(* IEC 61131-3 sources: guidance-for-physical-ai-production-designer-on-aws/source/plan2cell/crates/plan2cell/tests/fixtures/deploy_check/welding_cell_2_small/plc/codesys/head/GVL, 1 file *)

(* ---- GVL_Cell.st ---- *)
(*
 * GVL_Cell - generated by bt2plc 0.1.0 - DO NOT EDIT
 * Plan   : bt_1792076124_welding_cell_2_small (cell welding_cell_2_small)
 * Grants : planned ticket order
 * IL01   : R1#1 W03 > R2#2 W14 > R1#3 W06 > R2#4 W10 > R1#5 ROBOT1_S04 > R2#6 W12 > R1#7 W05 > R2#8 ROBOT2_S07 > R1#9 ROBOT1_S08 > R2#10 W07 > R1#11 HOME
 * IL02   : R2#1 W15 > R1#2 W02 > R2#3 W13 > R1#4 W01 > R2#5 W11 > R1#6 W04 > R2#7 ROBOT2_S06 > R1#8 W08 > R2#9 W09 > R1#10 ROBOT1_S09 > R2#11 HOME
 *)
{attribute 'qualified_only'}
VAR_GLOBAL CONSTANT
    (* ========================================================================
       DIMENSIONS (array bounds are literals; *_DIM >= 1)
       ======================================================================== *)
    N_ROBOTS                : INT := 2;
    N_ZONES                 : INT := 2;
    N_OPS                   : INT := 22;
    N_PREDS                 : INT := 0;

    (* ========================================================================
       PROTOCOL / TIMING
       ======================================================================== *)
    PLAN_ID                 : WORD := WORD#16#4F80;             (* fold of the plan fingerprint *)
    PROD_FOLGE              : WORD := WORD#11;                  (* default production Folge *)
    HOME_FOLGE              : WORD := WORD#125;                 (* blind homing *)
    JOB_NUMBER_BYTE         : BOOL := FALSE;                    (* FALSE: WORD LE bytes 2-3, TRUE: byte 2 *)
    PROFILE_VW              : BOOL := FALSE;                    (* TRUE: VW KS24 signal map and Folge handshake instead of the simulator telegram *)
    GRANT_POLICY            : E_GrantPolicy := E_GrantPolicy.GP_PLANNED;
    HOME_SEQUENTIAL         : BOOL := TRUE;
    AUTO_RUN                : BOOL := TRUE;                     (* start the next cycle automatically *)
    STEP_BYTE               : INT := 4;                         (* robot -> PLC, WORD LE op index *)
    REQ_BYTE                : INT := 28;                        (* robot -> PLC, DWORD LE zone requests *)
    GRANT_BYTE              : INT := 12;                        (* PLC -> robot, DWORD LE zone grants *)
    PLAN_ID_BYTE            : INT := 4;                         (* PLC -> robot, WORD LE plan id *)
    PERMIT_MASK             : DWORD := DWORD#16#80000000;       (* bit 31: permit predecessors *)
    T_RESET_PULSE           : TIME := T#1S;
    T_START_PULSE           : TIME := T#500MS;
    T_STOP_PULSE            : TIME := T#1S;
    T_HANDSHAKE             : TIME := T#5S;
    T_BRINGUP_LIMIT         : TIME := T#1M;                     (* safety enable: PROFINET connection set-up *)
    T_MISMATCH_DEBOUNCE     : TIME := T#200MS;
    T_STOP_DEBOUNCE         : TIME := T#200MS;                  (* job running: ProgRunning and ProgFinished low this long = robot stopped *)
    T_CYCLE_PAUSE           : TIME := T#2S;
    T_START_LIMIT           : TIME := T#15S;
    T_ABORT_LIMIT           : TIME := T#10S;
    T_HOME_LIMIT            : TIME := T#15S500MS;

    (* ========================================================================
       VW KS24 SIGNAL INDICES (used when PROFILE_VW; $IN/$OUT index, 1-based)
       ======================================================================== *)
    VW_READY_OUT            : INT := 9;                         (* O_R_Bereit *)
    VW_RK100_OUT            : INT := 10;                        (* O_R_RK100 safety circuit *)
    VW_AUTO_OUT             : INT := 12;                        (* O_R_Auto *)
    VW_ESTOP_OUT            : INT := 13;                        (* O_R_Notaus *)
    VW_END_OUT              : INT := 14;                        (* O_R_F_ENDE / LPKT *)
    VW_PF0_OUT              : INT := 15;                        (* O_R_PFO home position *)
    VW_STEP_OUT             : INT := 97;                        (* P_PktNr_SPS op index (16 bits) *)
    VW_REL_OUT              : INT := 41;                        (* interlock releases A41-56 *)
    VW_REQ_OUT              : INT := 81;                        (* interlock requests A81-96 *)
    VW_ERR_OUT              : INT := 225;                       (* VW_FEH_BIN_A error code (8 bits) *)
    VW_DRIVES_IN            : INT := 10;                        (* I_R_Ant_Ein *)
    VW_SRB_IN               : INT := 9;                         (* I_R_SRB Folge start *)
    VW_RESET_IN             : INT := 26;                        (* I_R_Quit_St acknowledge *)
    anInterlock             : ARRAY[1..4] OF INT := [0,0,0,0];  (* robot r, zone z -> VW interlock 1..16 (0 = not a member): index (r-1)*2+z *)

    (* ========================================================================
       ROBOTS (index = BT order)
       ======================================================================== *)
    asRobotTag              : ARRAY[1..2] OF STRING(16) := ['R1', 'R2'];
    asRobotNs               : ARRAY[1..2] OF STRING(32) := ['robot1', 'robot2'];
    abRobotActive           : ARRAY[1..2] OF BOOL := [TRUE, TRUE];
    abSafetyBypass          : ARRAY[1..2] OF BOOL := [TRUE, TRUE];(* SIMULATION ONLY: PROFIsafe slot-1 bits not required ([[robot]] safety_bypass) *)
    awRobotProdFolge        : ARRAY[1..2] OF WORD := [WORD#11, WORD#11];
    anRobotFirstOp          : ARRAY[1..2] OF INT := [1, 12];    (* op k of robot r: aOps[anRobotFirstOp[r] + k - 1] *)
    anRobotOpCount          : ARRAY[1..2] OF INT := [11, 11];

    (* ========================================================================
       ZONES - tickets of zone z: aTickets[anZoneFirst[z] .. anZoneFirst[z] + anZoneCount[z] - 1]
       ======================================================================== *)
    asZoneName              : ARRAY[1..2] OF STRING(8) := ['IL01', 'IL02'];
    anZoneFirst             : ARRAY[1..2] OF INT := [1, 12];
    anZoneCount             : ARRAY[1..2] OF INT := [11, 11];
    aTickets                : ARRAY[1..22] OF ST_Ticket := [
        (nRobot := 1, nOp := 1),    (* IL01 R1 #1 W03 *)
        (nRobot := 2, nOp := 2),    (* R2 #2 W14 *)
        (nRobot := 1, nOp := 3),    (* R1 #3 W06 *)
        (nRobot := 2, nOp := 4),    (* R2 #4 W10 *)
        (nRobot := 1, nOp := 5),    (* R1 #5 ROBOT1_S04 *)
        (nRobot := 2, nOp := 6),    (* R2 #6 W12 *)
        (nRobot := 1, nOp := 7),    (* R1 #7 W05 *)
        (nRobot := 2, nOp := 8),    (* R2 #8 ROBOT2_S07 *)
        (nRobot := 1, nOp := 9),    (* R1 #9 ROBOT1_S08 *)
        (nRobot := 2, nOp := 10),    (* R2 #10 W07 *)
        (nRobot := 1, nOp := 11),    (* R1 #11 HOME *)
        (nRobot := 2, nOp := 1),    (* IL02 R2 #1 W15 *)
        (nRobot := 1, nOp := 2),    (* R1 #2 W02 *)
        (nRobot := 2, nOp := 3),    (* R2 #3 W13 *)
        (nRobot := 1, nOp := 4),    (* R1 #4 W01 *)
        (nRobot := 2, nOp := 5),    (* R2 #5 W11 *)
        (nRobot := 1, nOp := 6),    (* R1 #6 W04 *)
        (nRobot := 2, nOp := 7),    (* R2 #7 ROBOT2_S06 *)
        (nRobot := 1, nOp := 8),    (* R1 #8 W08 *)
        (nRobot := 2, nOp := 9),    (* R2 #9 W09 *)
        (nRobot := 1, nOp := 10),    (* R1 #10 ROBOT1_S09 *)
        (nRobot := 2, nOp := 11)    (* R2 #11 HOME *)
    ];

    (* ========================================================================
       OPS - op k of robot r: aOps[anRobotFirstOp[r] + k - 1]
       ======================================================================== *)
    (* tLimit = 1.5 x tExpected + 5 s ; tZoneDeadline = 1.5 x ASAP grant + (5 + 0.2) s x depth + 10 s *)
    aOps                    : ARRAY[1..22] OF ST_OpInfo := [
        (nRobot := 1, nOp := 1, dwZoneMask := DWORD#16#00000001, nPredFirst := 0, nPredCount := 0, tExpected := T#3S409MS, tLimit := T#10S114MS, tZoneDeadline := T#10S, sName := 'W03'),    (* R1 #1 W03 *)
        (nRobot := 1, nOp := 2, dwZoneMask := DWORD#16#00000002, nPredFirst := 0, nPredCount := 0, tExpected := T#3S963MS, tLimit := T#10S945MS, tZoneDeadline := T#20S314MS, sName := 'W02'),    (* R1 #2 W02 *)
        (nRobot := 1, nOp := 3, dwZoneMask := DWORD#16#00000001, nPredFirst := 0, nPredCount := 0, tExpected := T#4S13MS, tLimit := T#11S20MS, tZoneDeadline := T#31S458MS, sName := 'W06'),    (* R1 #3 W06 *)
        (nRobot := 1, nOp := 4, dwZoneMask := DWORD#16#00000002, nPredFirst := 0, nPredCount := 0, tExpected := T#4S653MS, tLimit := T#11S980MS, tZoneDeadline := T#42S678MS, sName := 'W01'),    (* R1 #4 W01 *)
        (nRobot := 1, nOp := 5, dwZoneMask := DWORD#16#00000001, nPredFirst := 0, nPredCount := 0, tExpected := T#3S403MS, tLimit := T#10S105MS, tZoneDeadline := T#54S857MS, sName := 'ROBOT1_S04'),    (* R1 #5 ROBOT1_S04 *)
        (nRobot := 1, nOp := 6, dwZoneMask := DWORD#16#00000002, nPredFirst := 0, nPredCount := 0, tExpected := T#3S803MS, tLimit := T#10S705MS, tZoneDeadline := T#1M5S912MS, sName := 'W04'),    (* R1 #6 W04 *)
        (nRobot := 1, nOp := 7, dwZoneMask := DWORD#16#00000001, nPredFirst := 0, nPredCount := 0, tExpected := T#4S303MS, tLimit := T#11S455MS, tZoneDeadline := T#1M16S816MS, sName := 'W05'),    (* R1 #7 W05 *)
        (nRobot := 1, nOp := 8, dwZoneMask := DWORD#16#00000002, nPredFirst := 0, nPredCount := 0, tExpected := T#3S753MS, tLimit := T#10S630MS, tZoneDeadline := T#1M28S471MS, sName := 'W08'),    (* R1 #8 W08 *)
        (nRobot := 1, nOp := 9, dwZoneMask := DWORD#16#00000001, nPredFirst := 0, nPredCount := 0, tExpected := T#4S453MS, tLimit := T#11S680MS, tZoneDeadline := T#1M39S300MS, sName := 'ROBOT1_S08'),    (* R1 #9 ROBOT1_S08 *)
        (nRobot := 1, nOp := 10, dwZoneMask := DWORD#16#00000002, nPredFirst := 0, nPredCount := 0, tExpected := T#3S553MS, tLimit := T#10S330MS, tZoneDeadline := T#1M51S930MS, sName := 'ROBOT1_S09'),    (* R1 #10 ROBOT1_S09 *)
        (nRobot := 1, nOp := 11, dwZoneMask := DWORD#16#00000001, nPredFirst := 0, nPredCount := 0, tExpected := T#1S961MS, tLimit := T#7S942MS, tZoneDeadline := T#2M3S209MS, sName := 'HOME'),    (* R1 #11 HOME *)
        (nRobot := 2, nOp := 1, dwZoneMask := DWORD#16#00000002, nPredFirst := 0, nPredCount := 0, tExpected := T#3S409MS, tLimit := T#10S114MS, tZoneDeadline := T#10S, sName := 'W15'),    (* R2 #1 W15 *)
        (nRobot := 2, nOp := 2, dwZoneMask := DWORD#16#00000001, nPredFirst := 0, nPredCount := 0, tExpected := T#3S963MS, tLimit := T#10S945MS, tZoneDeadline := T#20S314MS, sName := 'W14'),    (* R2 #2 W14 *)
        (nRobot := 2, nOp := 3, dwZoneMask := DWORD#16#00000002, nPredFirst := 0, nPredCount := 0, tExpected := T#4S13MS, tLimit := T#11S20MS, tZoneDeadline := T#31S458MS, sName := 'W13'),    (* R2 #3 W13 *)
        (nRobot := 2, nOp := 4, dwZoneMask := DWORD#16#00000001, nPredFirst := 0, nPredCount := 0, tExpected := T#4S653MS, tLimit := T#11S980MS, tZoneDeadline := T#42S678MS, sName := 'W10'),    (* R2 #4 W10 *)
        (nRobot := 2, nOp := 5, dwZoneMask := DWORD#16#00000002, nPredFirst := 0, nPredCount := 0, tExpected := T#3S903MS, tLimit := T#10S855MS, tZoneDeadline := T#54S857MS, sName := 'W11'),    (* R2 #5 W11 *)
        (nRobot := 2, nOp := 6, dwZoneMask := DWORD#16#00000001, nPredFirst := 0, nPredCount := 0, tExpected := T#3S803MS, tLimit := T#10S705MS, tZoneDeadline := T#1M5S912MS, sName := 'W12'),    (* R2 #6 W12 *)
        (nRobot := 2, nOp := 7, dwZoneMask := DWORD#16#00000002, nPredFirst := 0, nPredCount := 0, tExpected := T#3S803MS, tLimit := T#10S705MS, tZoneDeadline := T#1M16S816MS, sName := 'ROBOT2_S06'),    (* R2 #7 ROBOT2_S06 *)
        (nRobot := 2, nOp := 8, dwZoneMask := DWORD#16#00000001, nPredFirst := 0, nPredCount := 0, tExpected := T#3S253MS, tLimit := T#9S880MS, tZoneDeadline := T#1M28S471MS, sName := 'ROBOT2_S07'),    (* R2 #8 ROBOT2_S07 *)
        (nRobot := 2, nOp := 9, dwZoneMask := DWORD#16#00000002, nPredFirst := 0, nPredCount := 0, tExpected := T#4S953MS, tLimit := T#12S430MS, tZoneDeadline := T#1M39S300MS, sName := 'W09'),    (* R2 #9 W09 *)
        (nRobot := 2, nOp := 10, dwZoneMask := DWORD#16#00000001, nPredFirst := 0, nPredCount := 0, tExpected := T#4S53MS, tLimit := T#11S80MS, tZoneDeadline := T#1M51S930MS, sName := 'W07'),    (* R2 #10 W07 *)
        (nRobot := 2, nOp := 11, dwZoneMask := DWORD#16#00000002, nPredFirst := 0, nPredCount := 0, tExpected := T#1S961MS, tLimit := T#7S942MS, tZoneDeadline := T#2M3S209MS, sName := 'HOME')    (* R2 #11 HOME *)
    ];

    (* ========================================================================
       PERMIT PREDECESSORS - op preds: aPreds[nPredFirst .. nPredFirst + nPredCount - 1]
       ======================================================================== *)
    aPreds                  : ARRAY[1..1] OF ST_Ticket := [
        (nRobot := 0, nOp := 0)    (* no permit predecessors *)
    ];
END_VAR
